(* PLC project g_trip_lockout_86_clean, Anonymous Benchmark Suite 1.0 *)
(* stored: creationDateTime 2026-09-02T00:00:00 *)

PROGRAM g_trip_lockout_86_clean
  VAR_INPUT
    protection_trip : BOOL;
    manual_reset : BOOL;
    reclose_request : BOOL;
    maint : BOOL;
  END_VAR
  VAR_OUTPUT
    lockout : BOOL;
    reclose : BOOL;
  END_VAR

(* LD diagram, written out as Structured Text *)
lockout := protection_trip OR lockout AND NOT manual_reset;
reclose := reclose_request AND NOT lockout AND NOT protection_trip;
END_PROGRAM

CONFIGURATION Config0
  RESOURCE Res0 ON PLC
    TASK tcyclic(INTERVAL := T#10ms, PRIORITY := 0);
    PROGRAM inst0 WITH tcyclic : g_trip_lockout_86_clean;
  END_RESOURCE
END_CONFIGURATION
